Universal Robots URScript: T007_mistralai_Devstral-Small-2-24B-Instruct-2512_edit_perf_rep1.urscript

# Task: T007 — Curved contour weld — hybrid mode
# Optimized for faster cycle time
# Operating mode: hybrid | Max TCP speed: 0.300 m/s
# Robot: ur5e

def task_T007():
  TCP_SPEED_CAP = 0.300
  def safe_movel(pose, a, v, r):
    if (v > TCP_SPEED_CAP):
      popup("TCP speed cap exceeded", error=True)
      halt
    end
    movel(pose, a=a, v=v, r=r)
  end

  # [1] Home position (faster acceleration)
  movej([0.0000, -1.5708, 1.5708, -1.5708, -1.5708, 0.0000], a=1.5700, v=0.7500)

  # [2] Approach above weld fixture (faster)
  safe_movel(p[0.450000, 0.000000, 0.350000, 0.0000, 3.1416, 0.0000], 1.2000, 0.2500, 0.0100)

  # [3] Descend to weld start (faster)
  safe_movel(p[0.450000, 0.000000, 0.200000, 0.0000, 3.1416, 0.0000], 0.7000, 0.1000, 0.0010)

  # [4] Gas pre-flow ON
  set_digital_out(1, True)

  # [5] Gas stabilization (reduced time)
  sleep(0.3000)

  # [6] Arc ON
  set_digital_out(0, True)
  set_analog_out(0, 0.500)
  set_analog_out(1, 0.400)

  # [7] Weld midpoint (faster)
  safe_movel(p[0.550000, 0.150000, 0.200000, 0.0000, 3.1416, 0.0000], 0.3000, 0.0600, 0.0050)

  # [8] Weld end (faster)
  safe_movel(p[0.500000, 0.300000, 0.200000, 0.0000, 3.1416, 0.0000], 0.3000, 0.0600, 0.0)

  # [9] Arc OFF
  set_digital_out(0, False)
  set_analog_out(0, 0.0)
  set_analog_out(1, 0.0)

  # [10] Post-weld gas flow (reduced time)
  sleep(0.5000)

  # [11] Gas flow OFF
  set_digital_out(1, False)

  # [12] Retract above weld end (faster)
  safe_movel(p[0.500000, 0.300000, 0.380000, 0.0000, 3.1416, 0.0000], 1.2000, 0.2500, 0.0100)

  # [13] Return to home (faster acceleration)
  movej([0.0000, -1.5708, 1.5708, -1.5708, -1.5708, 0.0000], a=1.5700, v=0.7500)

end

# Entry point
task_T007()
